(* Logix 5000 project; controller CIP_14485201 vendor 1 type 14 code 216 rev 38.11; software revision 38.01; part 6 of 12 *)
(* tags used below, declared in another part *)
   Alarm_Ack : INT[8];   // ALARMS ACKNOWLEDGE BITS
   Alarm_Ack_All_PB : BOOL;   // SYSTEM ALARM ACK ALL PUSHBUTTON ON ALARM PAGE
   Alarm_Present : INT[8];   // ALARM MSGS 1-127 PRESENT BITS
   Alarm_Remote_Ack_All : BOOL;   // SYSTEM ALARM ACK ALL TAG USED ON ALARM SETUP ADVANCED TAB TOGGLES EVEYTIME THE ACK_ALL BUTTON IS PUSHED
   Alarm_Status_Reset : BOOL;   // SYSTEM ALARM ACK ALL TAG USED ON ALARM SETUP ADVANCED TAB TOGGLES EVERYTIME THE HISTORY CLEAR ALL IS PUSHED
   Bit : BOOL[128];   // BIT
   One_Shot : BOOL[128];   // ONE SHOT ARRAY
   Panelview : INT[40];   // PANELVIEW CONTROL
   SYS_Bit : BOOL[128];   // SYSTEM BIT
   SYS_Timer : TIMER[60];   // SYSTEM TIMER
(* MainProgram, continued *)

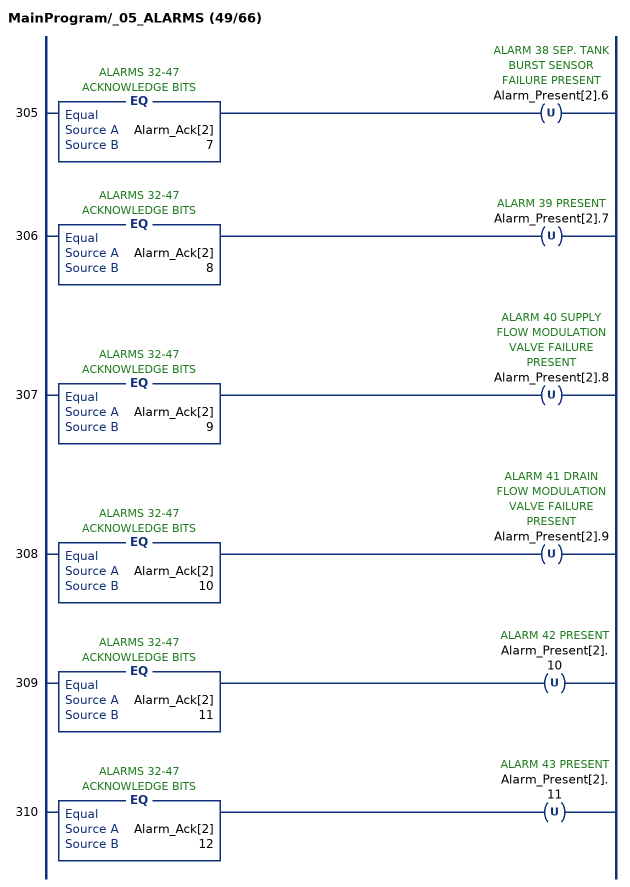
   [picture p76: MainProgram/_05_ALARMS rungs 305-310]
   305: EQ(Alarm_Ack[2],7)OTU(Alarm_Present[2].6);
   306: EQ(Alarm_Ack[2],8)OTU(Alarm_Present[2].7);
   307: EQ(Alarm_Ack[2],9)OTU(Alarm_Present[2].8);
   308: EQ(Alarm_Ack[2],10)OTU(Alarm_Present[2].9);
   309: EQ(Alarm_Ack[2],11)OTU(Alarm_Present[2].10);
   310: EQ(Alarm_Ack[2],12)OTU(Alarm_Present[2].11);
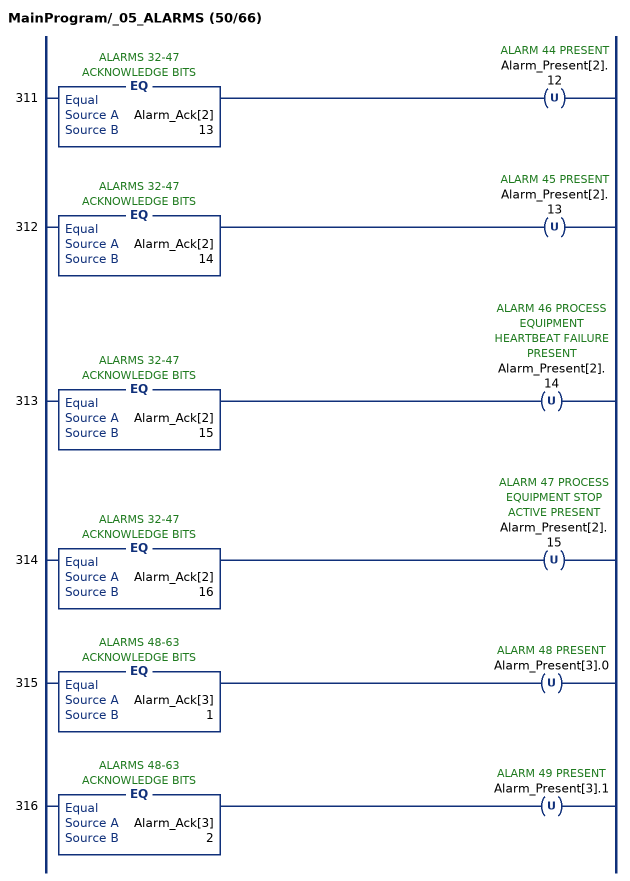
   311: EQ(Alarm_Ack[2],13)OTU(Alarm_Present[2].12);
   312: EQ(Alarm_Ack[2],14)OTU(Alarm_Present[2].13);
   313: EQ(Alarm_Ack[2],15)OTU(Alarm_Present[2].14);
   314: EQ(Alarm_Ack[2],16)OTU(Alarm_Present[2].15);
   315: EQ(Alarm_Ack[3],1)OTU(Alarm_Present[3].0);
   316: EQ(Alarm_Ack[3],2)OTU(Alarm_Present[3].1);
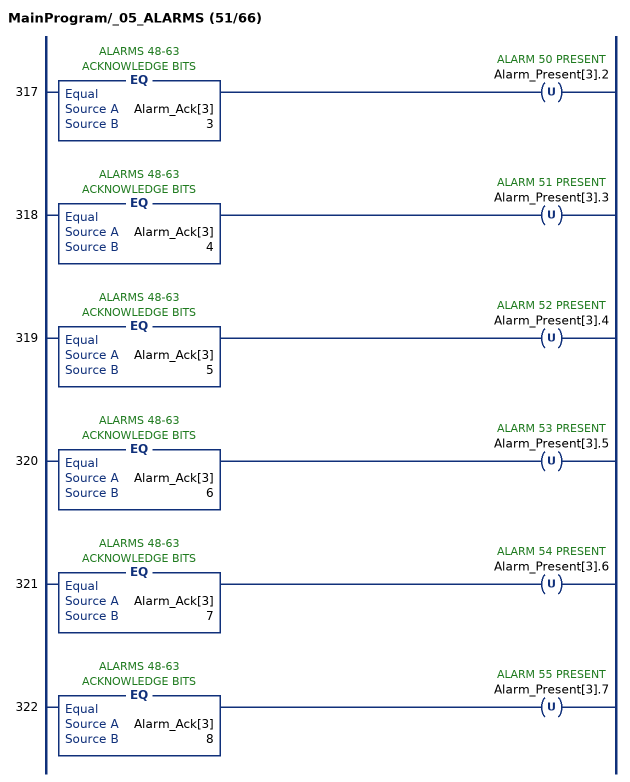
   317: EQ(Alarm_Ack[3],3)OTU(Alarm_Present[3].2);
   318: EQ(Alarm_Ack[3],4)OTU(Alarm_Present[3].3);
   319: EQ(Alarm_Ack[3],5)OTU(Alarm_Present[3].4);
   320: EQ(Alarm_Ack[3],6)OTU(Alarm_Present[3].5);
   321: EQ(Alarm_Ack[3],7)OTU(Alarm_Present[3].6);
   322: EQ(Alarm_Ack[3],8)OTU(Alarm_Present[3].7);
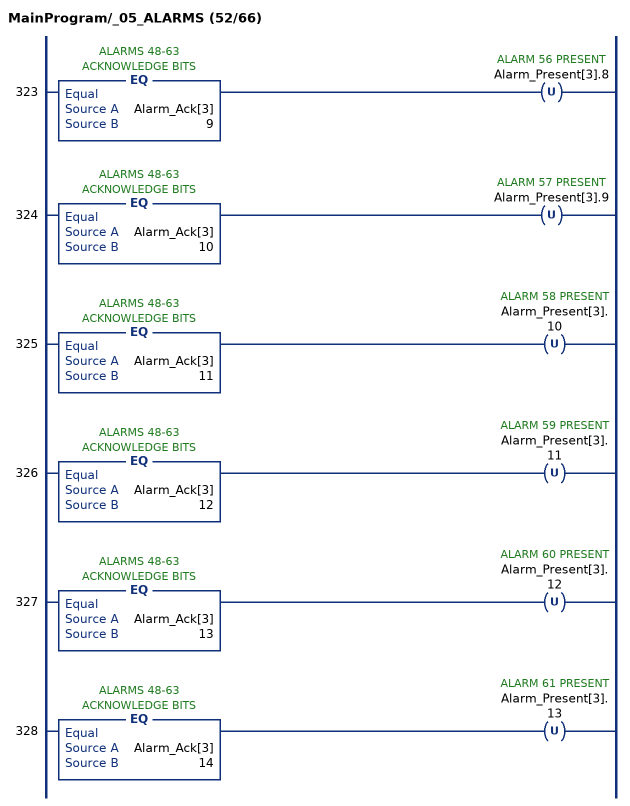
   323: EQ(Alarm_Ack[3],9)OTU(Alarm_Present[3].8);
   324: EQ(Alarm_Ack[3],10)OTU(Alarm_Present[3].9);
   325: EQ(Alarm_Ack[3],11)OTU(Alarm_Present[3].10);
   326: EQ(Alarm_Ack[3],12)OTU(Alarm_Present[3].11);
   327: EQ(Alarm_Ack[3],13)OTU(Alarm_Present[3].12);
   328: EQ(Alarm_Ack[3],14)OTU(Alarm_Present[3].13);
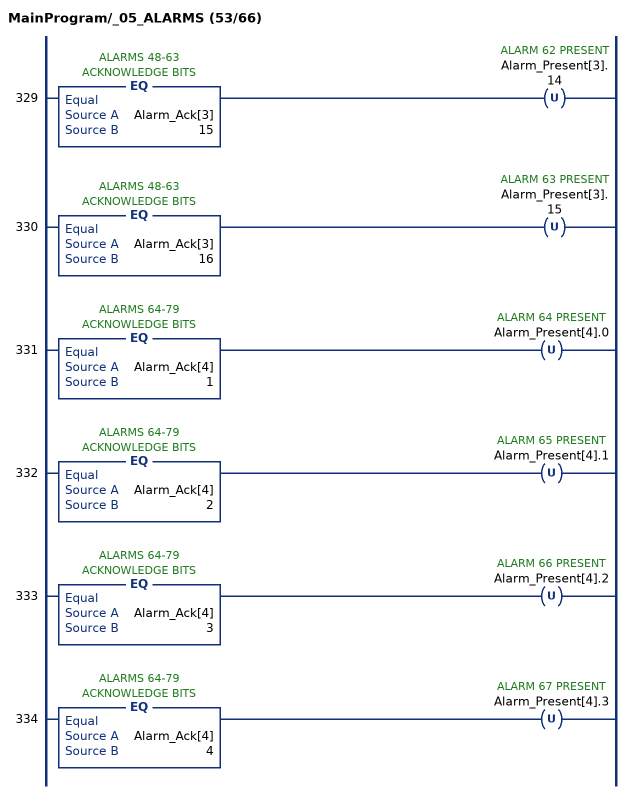
   329: EQ(Alarm_Ack[3],15)OTU(Alarm_Present[3].14);
   330: EQ(Alarm_Ack[3],16)OTU(Alarm_Present[3].15);
   331: EQ(Alarm_Ack[4],1)OTU(Alarm_Present[4].0);
   332: EQ(Alarm_Ack[4],2)OTU(Alarm_Present[4].1);
   333: EQ(Alarm_Ack[4],3)OTU(Alarm_Present[4].2);
   334: EQ(Alarm_Ack[4],4)OTU(Alarm_Present[4].3);
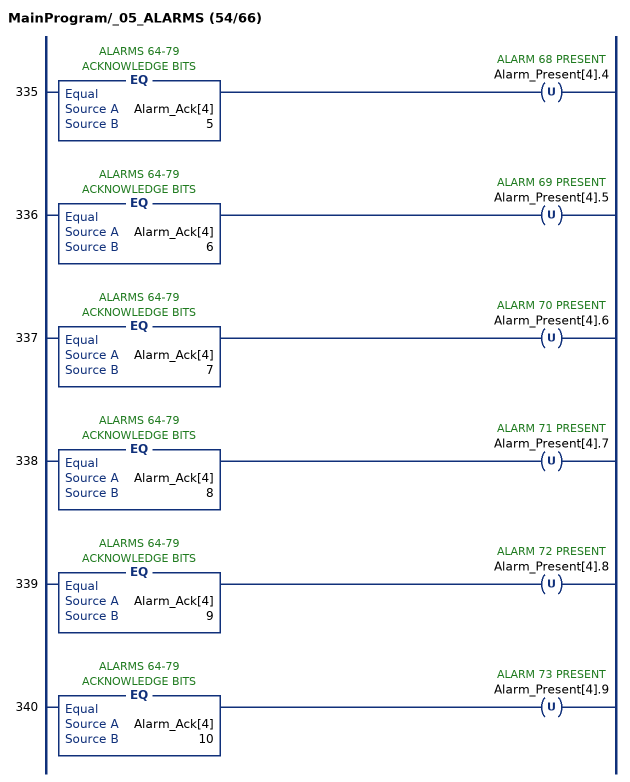
   335: EQ(Alarm_Ack[4],5)OTU(Alarm_Present[4].4);
   336: EQ(Alarm_Ack[4],6)OTU(Alarm_Present[4].5);
   337: EQ(Alarm_Ack[4],7)OTU(Alarm_Present[4].6);
   338: EQ(Alarm_Ack[4],8)OTU(Alarm_Present[4].7);
   339: EQ(Alarm_Ack[4],9)OTU(Alarm_Present[4].8);
   340: EQ(Alarm_Ack[4],10)OTU(Alarm_Present[4].9);
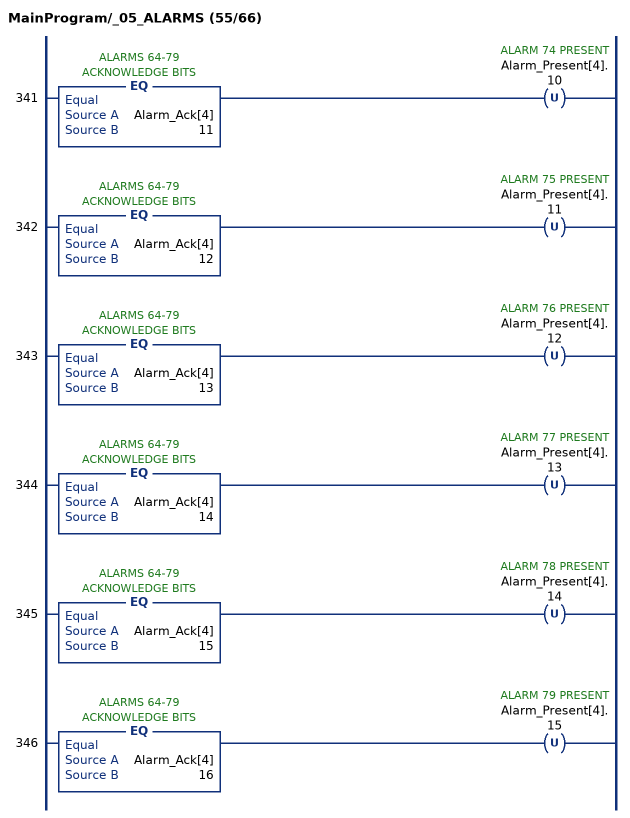
   341: EQ(Alarm_Ack[4],11)OTU(Alarm_Present[4].10);
   342: EQ(Alarm_Ack[4],12)OTU(Alarm_Present[4].11);
   343: EQ(Alarm_Ack[4],13)OTU(Alarm_Present[4].12);
   344: EQ(Alarm_Ack[4],14)OTU(Alarm_Present[4].13);
   345: EQ(Alarm_Ack[4],15)OTU(Alarm_Present[4].14);
   346: EQ(Alarm_Ack[4],16)OTU(Alarm_Present[4].15);
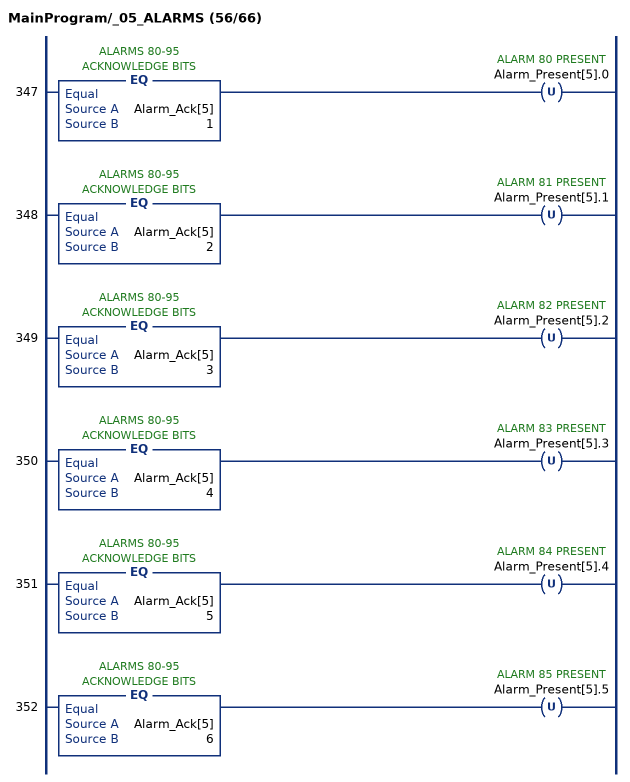
   347: EQ(Alarm_Ack[5],1)OTU(Alarm_Present[5].0);
   348: EQ(Alarm_Ack[5],2)OTU(Alarm_Present[5].1);
   349: EQ(Alarm_Ack[5],3)OTU(Alarm_Present[5].2);
   350: EQ(Alarm_Ack[5],4)OTU(Alarm_Present[5].3);
   351: EQ(Alarm_Ack[5],5)OTU(Alarm_Present[5].4);
   352: EQ(Alarm_Ack[5],6)OTU(Alarm_Present[5].5);
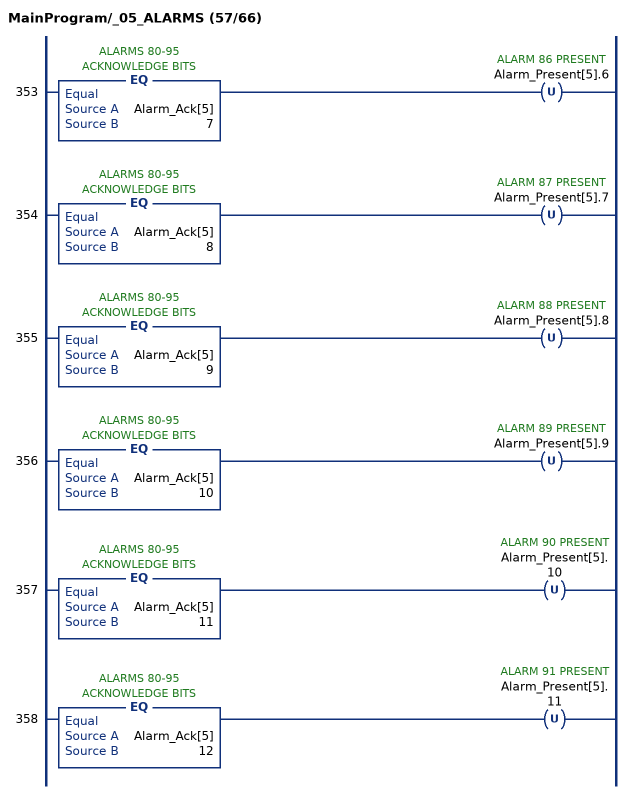
   353: EQ(Alarm_Ack[5],7)OTU(Alarm_Present[5].6);
   354: EQ(Alarm_Ack[5],8)OTU(Alarm_Present[5].7);
   355: EQ(Alarm_Ack[5],9)OTU(Alarm_Present[5].8);
   356: EQ(Alarm_Ack[5],10)OTU(Alarm_Present[5].9);
   357: EQ(Alarm_Ack[5],11)OTU(Alarm_Present[5].10);
   358: EQ(Alarm_Ack[5],12)OTU(Alarm_Present[5].11);
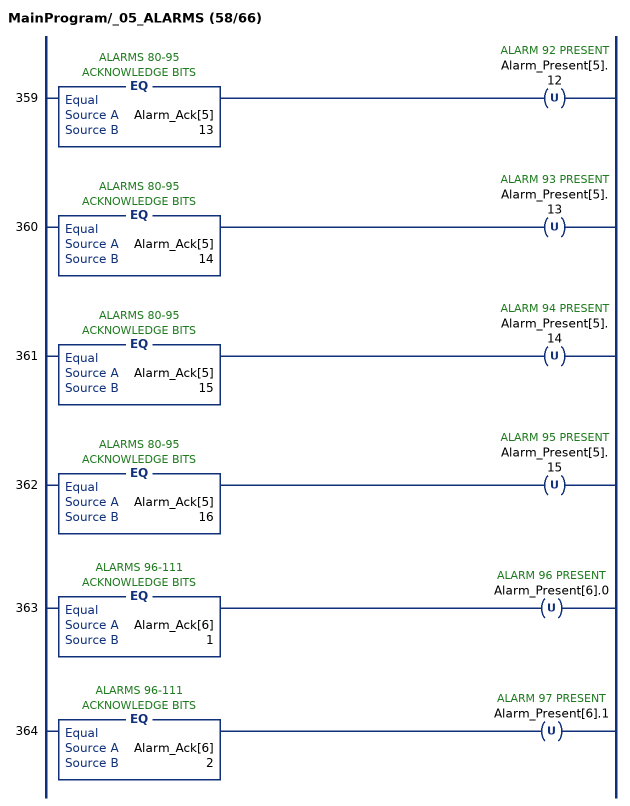
   359: EQ(Alarm_Ack[5],13)OTU(Alarm_Present[5].12);
   360: EQ(Alarm_Ack[5],14)OTU(Alarm_Present[5].13);
   361: EQ(Alarm_Ack[5],15)OTU(Alarm_Present[5].14);
   362: EQ(Alarm_Ack[5],16)OTU(Alarm_Present[5].15);
   363: EQ(Alarm_Ack[6],1)OTU(Alarm_Present[6].0);
   364: EQ(Alarm_Ack[6],2)OTU(Alarm_Present[6].1);
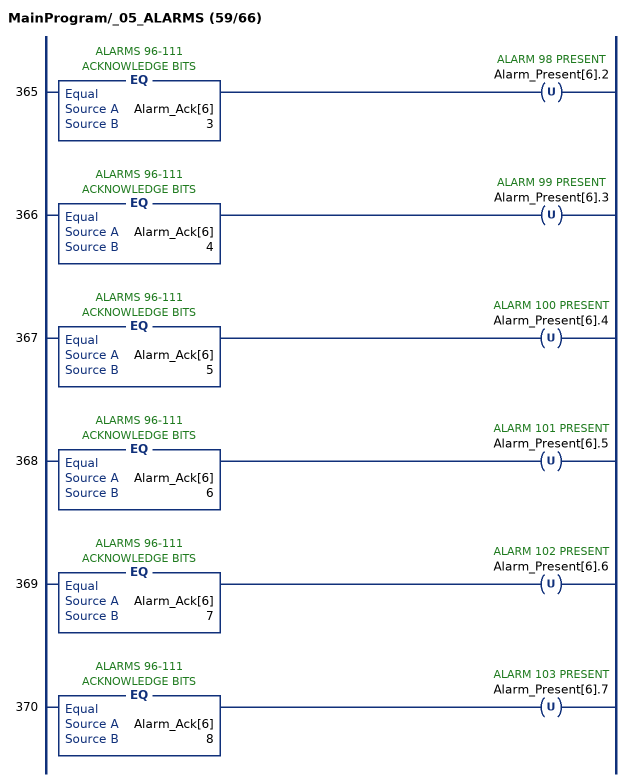
   365: EQ(Alarm_Ack[6],3)OTU(Alarm_Present[6].2);
   366: EQ(Alarm_Ack[6],4)OTU(Alarm_Present[6].3);
   367: EQ(Alarm_Ack[6],5)OTU(Alarm_Present[6].4);
   368: EQ(Alarm_Ack[6],6)OTU(Alarm_Present[6].5);
   369: EQ(Alarm_Ack[6],7)OTU(Alarm_Present[6].6);
   370: EQ(Alarm_Ack[6],8)OTU(Alarm_Present[6].7);
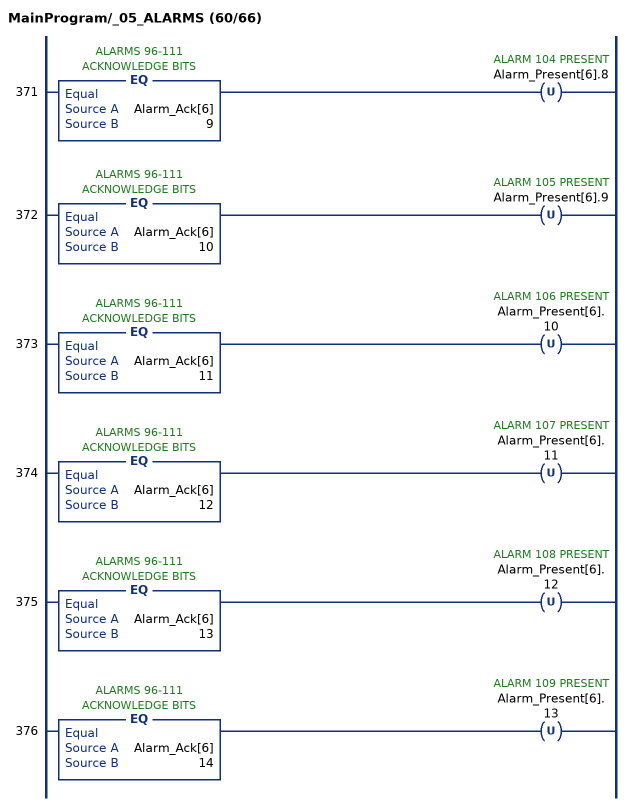
   371: EQ(Alarm_Ack[6],9)OTU(Alarm_Present[6].8);
   372: EQ(Alarm_Ack[6],10)OTU(Alarm_Present[6].9);
   373: EQ(Alarm_Ack[6],11)OTU(Alarm_Present[6].10);
   374: EQ(Alarm_Ack[6],12)OTU(Alarm_Present[6].11);
   375: EQ(Alarm_Ack[6],13)OTU(Alarm_Present[6].12);
   376: EQ(Alarm_Ack[6],14)OTU(Alarm_Present[6].13);
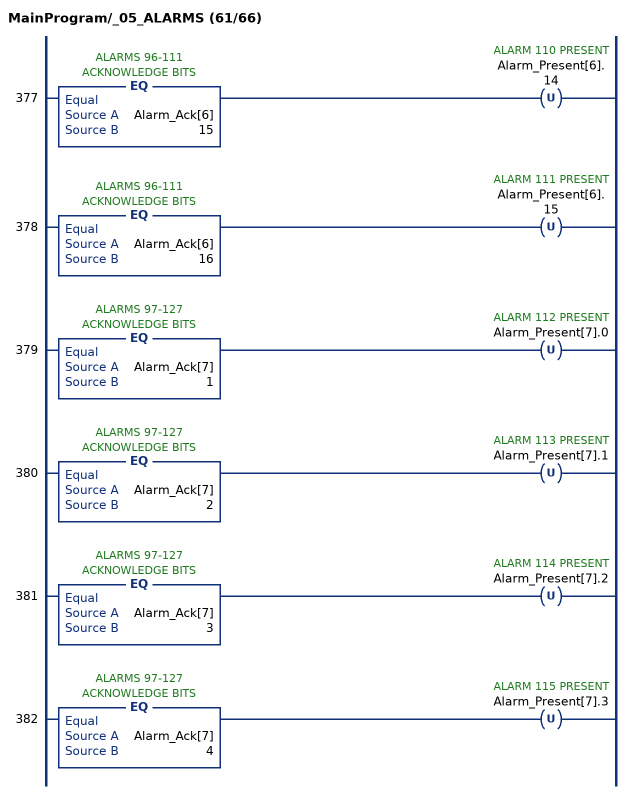
   377: EQ(Alarm_Ack[6],15)OTU(Alarm_Present[6].14);
   378: EQ(Alarm_Ack[6],16)OTU(Alarm_Present[6].15);
   379: EQ(Alarm_Ack[7],1)OTU(Alarm_Present[7].0);
   380: EQ(Alarm_Ack[7],2)OTU(Alarm_Present[7].1);
   381: EQ(Alarm_Ack[7],3)OTU(Alarm_Present[7].2);
   382: EQ(Alarm_Ack[7],4)OTU(Alarm_Present[7].3);
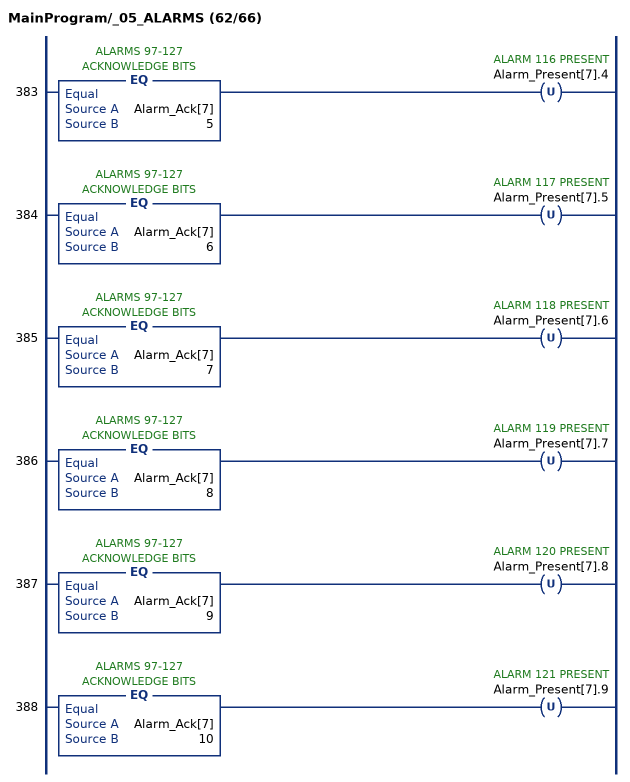
   383: EQ(Alarm_Ack[7],5)OTU(Alarm_Present[7].4);
   384: EQ(Alarm_Ack[7],6)OTU(Alarm_Present[7].5);
   385: EQ(Alarm_Ack[7],7)OTU(Alarm_Present[7].6);
   386: EQ(Alarm_Ack[7],8)OTU(Alarm_Present[7].7);
   387: EQ(Alarm_Ack[7],9)OTU(Alarm_Present[7].8);
   388: EQ(Alarm_Ack[7],10)OTU(Alarm_Present[7].9);
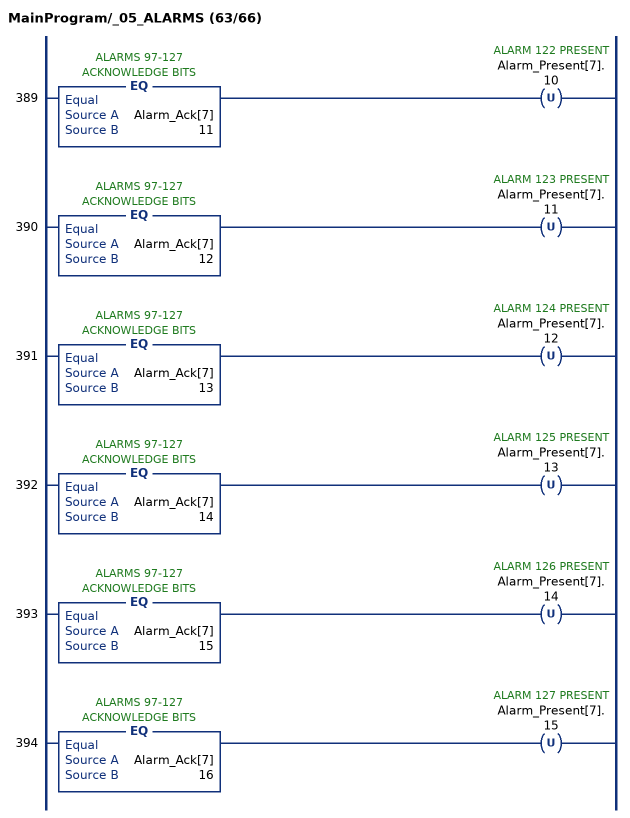
   389: EQ(Alarm_Ack[7],11)OTU(Alarm_Present[7].10);
   390: EQ(Alarm_Ack[7],12)OTU(Alarm_Present[7].11);
   391: EQ(Alarm_Ack[7],13)OTU(Alarm_Present[7].12);
   392: EQ(Alarm_Ack[7],14)OTU(Alarm_Present[7].13);
   393: EQ(Alarm_Ack[7],15)OTU(Alarm_Present[7].14);
   394: EQ(Alarm_Ack[7],16)OTU(Alarm_Present[7].15);
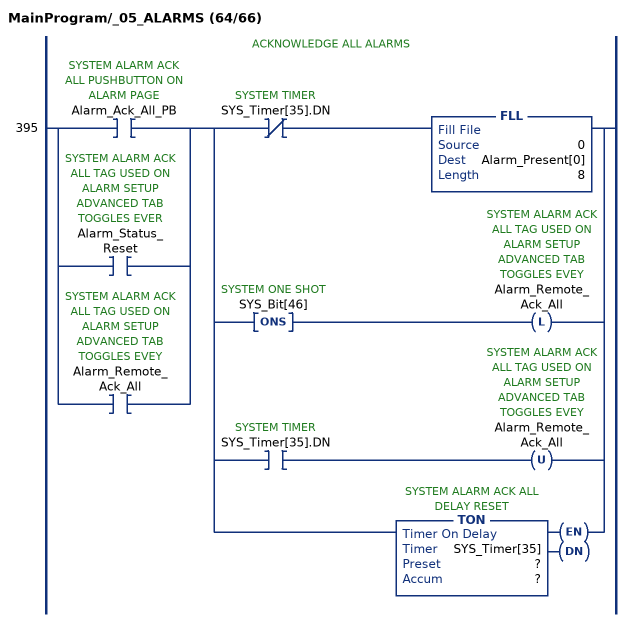
   // ACKNOWLEDGE ALL ALARMS
   395: [XIC(Alarm_Ack_All_PB) ,XIC(Alarm_Status_Reset) ,XIC(Alarm_Remote_Ack_All) ][XIO(SYS_Timer[35].DN) FLL(0,Alarm_Present[0],8) ,ONS(SYS_Bit[46]) OTL(Alarm_Remote_Ack_All) ,XIC(SYS_Timer[35].DN) OTU(Alarm_Remote_Ack_All) ,TON(SYS_Timer[35],?,?) ];
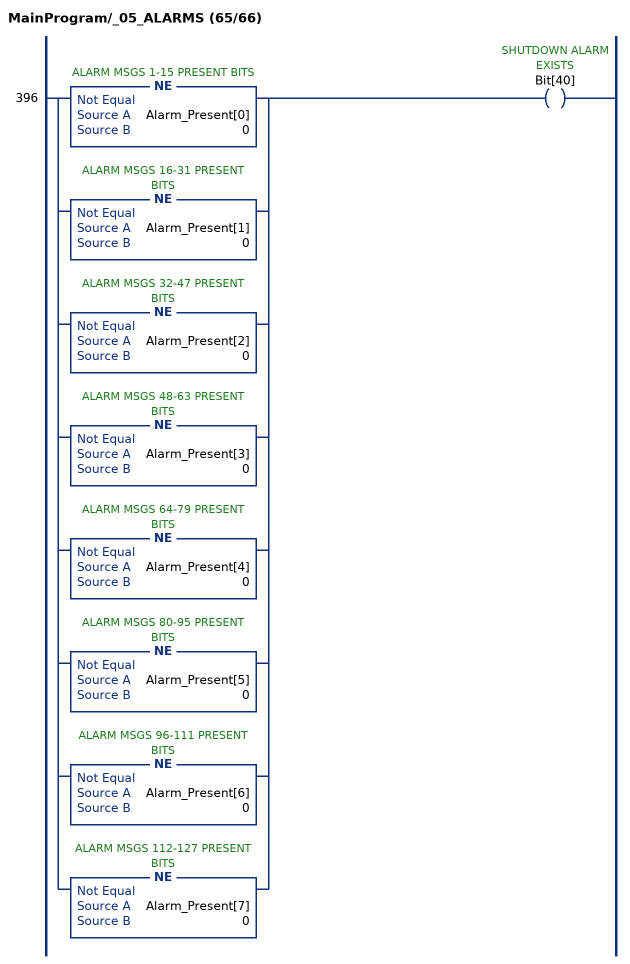
   396: [NE(Alarm_Present[0],0) ,NE(Alarm_Present[1],0) ,NE(Alarm_Present[2],0) ,NE(Alarm_Present[3],0) ,NE(Alarm_Present[4],0) ,NE(Alarm_Present[5],0) ,NE(Alarm_Present[6],0) ,NE(Alarm_Present[7],0) ]OTE(Bit[40]);
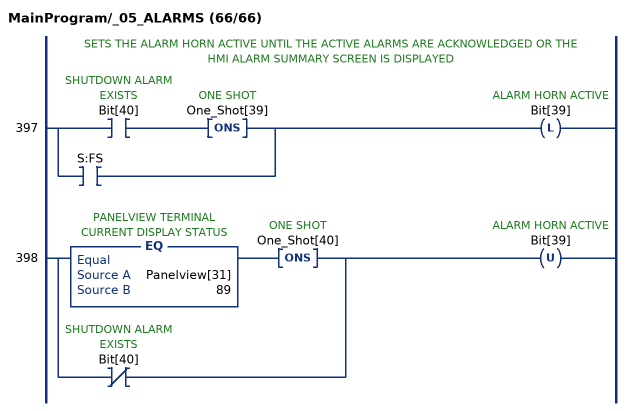
   // SETS THE ALARM HORN ACTIVE UNTIL THE ACTIVE ALARMS ARE ACKNOWLEDGED OR THE HMI ALARM SUMMARY SCREEN IS DISPLAYED
   397: [XIC(Bit[40]) ONS(One_Shot[39]) ,XIC(S:FS) ]OTL(Bit[39]);
   398: [EQ(Panelview[31],89) ONS(One_Shot[40]) ,XIO(Bit[40]) ]OTU(Bit[39]);
END_ROUTINE
